(* IEC 61131-3 sources: AI_Prediciton_FInder_Energy_meter/plc/src, 8 files *)

(* ---- U_Word32.st ---- *)
// DUT (UNION) - reinterprets 32 bits as DWORD, REAL or DINT
TYPE U_Word32 :
UNION
    dwRaw : DWORD;
    rReal : REAL;
    diInt : DINT;
END_UNION
END_TYPE

(* ---- GVL_Meter.st ---- *)
// GVL - raw Modbus channels and Modbus TCP input registers
VAR_GLOBAL
    // Finder 7M.24 #1 (Modbus RTU address 2) - mapped in Modbus_Server_COM_Port I/O Mapping
    awFinder1Power      : ARRAY[0..11] OF WORD;  // 32490..32501: Pt, Qt, St, PFt, f, U1 (REAL, high word first)
    awFinder1Current    : ARRAY[0..1] OF WORD;   // 32516..32517: I1 (REAL)
    awFinder1EnergyExp  : ARRAY[0..3] OF WORD;   // 30401..30404: exponents n1..n4 (INT)
    awFinder1EnergyMant : ARRAY[0..7] OF WORD;   // 30406..30413: mantissas n1..n4 (DINT, high word first)
    awFinder1Identity   : ARRAY[0..11] OF WORD;  // 30001..30012: model (0..7) + serial (8..11), ASCII
    awFinder1MaxRegs    : ARRAY[0..0] OF WORD;   // 30099: max registers per request
    // E2-PLC2 (25.11.2026): new channels, existing ones unchanged
    awFinder1Quality    : ARRAY[0..25] OF WORD;  // 32570..32595: angle U1-I1 [0..1], THD I1 [18..19], THD U1 [24..25] (REAL)
    awFinder1Temp       : ARRAY[0..1] OF WORD;   // 32658..32659: internal temperature (REAL, degC)
    awFinder1RunTime    : ARRAY[0..1] OF WORD;   // 32480..32481: run time (REAL, s - type to be confirmed)

    // Modbus TCP server input registers (FC04) - mapped in ModbusTCP_Server_Device I/O Mapping
    awTcpInputRegs      : ARRAY[0..99] OF WORD;
END_VAR

(* ---- FC_PutDword.st ---- *)
// FUNCTION, return type BOOL - writes 32 bits into two registers, high word first
FUNCTION FC_PutDword : BOOL
VAR_IN_OUT
    awRegs : ARRAY[0..99] OF WORD;
END_VAR
VAR_INPUT
    iIndex  : INT;    // index of the first (high) register
    dwValue : DWORD;
END_VAR
// --- code ---
IF (iIndex < 0) OR (iIndex > 98) THEN
    FC_PutDword := FALSE;
    RETURN;
END_IF
awRegs[iIndex]     := DWORD_TO_WORD(SHR(dwValue, 16));
awRegs[iIndex + 1] := DWORD_TO_WORD(dwValue);
FC_PutDword := TRUE;

(* ---- FC_PutReal.st ---- *)
// FUNCTION, return type BOOL - writes REAL (IEEE 754) into two registers, high word first
FUNCTION FC_PutReal : BOOL
VAR_IN_OUT
    awRegs : ARRAY[0..99] OF WORD;
END_VAR
VAR_INPUT
    iIndex : INT;
    rValue : REAL;
END_VAR
VAR
    uConv : U_Word32;
END_VAR
// --- code ---
uConv.rReal := rValue;
FC_PutReal := FC_PutDword(awRegs := awRegs, iIndex := iIndex, dwValue := uConv.dwRaw);

(* ---- FC_WordsToDword.st ---- *)
// FUNCTION, return type DWORD
FUNCTION FC_WordsToDword : DWORD
VAR_INPUT
    wFirst     : WORD;  // register with lower address
    wSecond    : WORD;  // register with higher address
    xSwapWords : BOOL;  // FALSE = first register is the high word (Finder 7M.24, verified 23.11.2026)
END_VAR
// --- code ---
IF xSwapWords THEN
    FC_WordsToDword := SHL(WORD_TO_DWORD(wSecond), 16) OR WORD_TO_DWORD(wFirst);
ELSE
    FC_WordsToDword := SHL(WORD_TO_DWORD(wFirst), 16) OR WORD_TO_DWORD(wSecond);
END_IF

(* ---- FC_WordsToReal.st ---- *)
// FUNCTION, return type REAL
FUNCTION FC_WordsToReal : REAL
VAR_INPUT
    wFirst     : WORD;
    wSecond    : WORD;
    xSwapWords : BOOL;
END_VAR
VAR
    uConv : U_Word32;
END_VAR
// --- code ---
uConv.dwRaw := FC_WordsToDword(wFirst := wFirst, wSecond := wSecond, xSwapWords := xSwapWords);
FC_WordsToReal := uConv.rReal;

(* ---- FB_EnergyMeter.st ---- *)
// FUNCTION_BLOCK - one instance = one Finder 7M.24 meter
FUNCTION_BLOCK FB_EnergyMeter
VAR_INPUT
    xCommError        : BOOL;                   // <device>.xError of the Modbus server (COM) instance
    uiModbusErrorCode : UINT;                   // <device>.byModbusError (MB_ErrorCodes)
    awPower           : ARRAY[0..11] OF WORD;
    awCurrent         : ARRAY[0..1] OF WORD;
    awEnergyExp       : ARRAY[0..3] OF WORD;
    awEnergyMant      : ARRAY[0..7] OF WORD;
    awIdentity        : ARRAY[0..11] OF WORD;
    awQuality         : ARRAY[0..25] OF WORD;   // 32570..32595 (map v2, 25.11.2026)
    awTemp            : ARRAY[0..1] OF WORD;    // 32658..32659
    awRunTime         : ARRAY[0..1] OF WORD;    // 32480..32481
    xSwapWords        : BOOL := FALSE;          // Finder 7M.24: high word first -> FALSE
    tErrorHold        : TIME := T#3S;           // COMM_ERROR is cleared only after this time without any error
END_VAR
VAR_OUTPUT
    rActivePower_W     : REAL;
    rReactivePower_var : REAL;
    rApparentPower_VA  : REAL;
    rPowerFactor       : REAL;
    rFrequency_Hz      : REAL;
    rVoltage_V         : REAL;
    rCurrent_A         : REAL;
    diEnergyImportMant : DINT;   // n1, Wh = mant * 10^exp
    iEnergyImportExp   : INT;
    diEnergyExportMant : DINT;   // n3
    iEnergyExportExp   : INT;
    rEnergyImport_kWh  : REAL;
    rEnergyExport_kWh  : REAL;
    diReactivePosMant  : DINT;   // n2 (energy at Q > 0), varh = mant * 10^exp
    iReactivePosExp    : INT;
    diReactiveNegMant  : DINT;   // n4 (energy at Q < 0)
    iReactiveNegExp    : INT;
    rThdVoltage_pct    : REAL;   // THD U1, 32594
    rThdCurrent_pct    : REAL;   // THD I1, 32588
    rPhaseAngle_deg    : REAL;   // angle U1-I1, 32570 (negative at Q < 0, measured 25.11.2026)
    rTemperature_C     : REAL;   // internal meter temperature, 32658
    rRunTime_s         : REAL;   // meter run time, 32480
    awSerial           : ARRAY[0..3] OF WORD;
    sSerial            : STRING(8);
    uiStatus           : UINT;   // 0 = OK, 1 = COMM_ERROR, 2 = NO_DATA (no answer since start)
    uiErrorCode        : UINT;   // last non-zero MB_ErrorCodes value while not OK, 0 when OK
    uiErrorCount       : UINT;   // number of communication outages since start (wraps at 65535)
    udiDataAge_ms      : UDINT;  // 0 when OK; time since last confirmed OK state otherwise
END_VAR
VAR CONSTANT
    STATUS_OK         : UINT := 0;
    STATUS_COMM_ERROR : UINT := 1;
    STATUS_NO_DATA    : UINT := 2;
END_VAR
VAR
    xErrorSeen       : BOOL;   // at least one raw error since start
    xErrorActive     : BOOL;   // debounced error: raw error within the last tErrorHold
    xErrorActivePrev : BOOL;
    xDataSeen        : BOOL;
    tNow             : TIME;
    tLastOk          : TIME;
    tLastErr         : TIME;
    uiLastErrCode    : UINT;
    uConv            : U_Word32;
    pbySerial        : POINTER TO BYTE;
    i                : INT;
END_VAR
// --- code ---
// 1. Communication status (debounced: xError of the COM device drops between transactions;
//    fixed 23.11.2026 after checklist test 5)
tNow := TIME();
IF xCommError THEN
    xErrorSeen := TRUE;
    tLastErr   := tNow;
    IF uiModbusErrorCode <> 0 THEN
        uiLastErrCode := uiModbusErrorCode;
    END_IF
END_IF

xErrorActive := xErrorSeen AND ((tNow - tLastErr) < tErrorHold);

IF NOT xErrorActive THEN
    tLastOk := tNow;
END_IF
IF xErrorActive AND NOT xErrorActivePrev THEN
    uiErrorCount := uiErrorCount + 1;            // one outage = one count
END_IF
xErrorActivePrev := xErrorActive;

// Meter has answered at least once when the serial number registers are not zero
IF (awIdentity[8] <> 0) OR (awIdentity[9] <> 0) THEN
    xDataSeen := TRUE;
END_IF

IF NOT xDataSeen THEN
    uiStatus      := STATUS_NO_DATA;
    uiErrorCode   := uiLastErrCode;
    udiDataAge_ms := 16#FFFFFFFF;
ELSIF xErrorActive THEN
    uiStatus      := STATUS_COMM_ERROR;
    uiErrorCode   := uiLastErrCode;
    udiDataAge_ms := TIME_TO_UDINT(tNow - tLastOk);
ELSE
    uiStatus      := STATUS_OK;
    uiErrorCode   := 0;
    uiLastErrCode := 0;
    udiDataAge_ms := 0;
END_IF

// 2. Instantaneous values (IEEE 754 block 32490..32501, 32516)
rActivePower_W     := FC_WordsToReal(wFirst := awPower[0],  wSecond := awPower[1],  xSwapWords := xSwapWords);
rReactivePower_var := FC_WordsToReal(wFirst := awPower[2],  wSecond := awPower[3],  xSwapWords := xSwapWords);
rApparentPower_VA  := FC_WordsToReal(wFirst := awPower[4],  wSecond := awPower[5],  xSwapWords := xSwapWords);
rPowerFactor       := FC_WordsToReal(wFirst := awPower[6],  wSecond := awPower[7],  xSwapWords := xSwapWords);
rFrequency_Hz      := FC_WordsToReal(wFirst := awPower[8],  wSecond := awPower[9],  xSwapWords := xSwapWords);
rVoltage_V         := FC_WordsToReal(wFirst := awPower[10], wSecond := awPower[11], xSwapWords := xSwapWords);
rCurrent_A         := FC_WordsToReal(wFirst := awCurrent[0], wSecond := awCurrent[1], xSwapWords := xSwapWords);

// 3. Energy counters: Wh = mantissa * 10^exponent (n1 = import, n3 = export - to confirm on display)
uConv.dwRaw := FC_WordsToDword(wFirst := awEnergyMant[0], wSecond := awEnergyMant[1], xSwapWords := xSwapWords);
diEnergyImportMant := uConv.diInt;
iEnergyImportExp   := WORD_TO_INT(awEnergyExp[0]);

uConv.dwRaw := FC_WordsToDword(wFirst := awEnergyMant[4], wSecond := awEnergyMant[5], xSwapWords := xSwapWords);
diEnergyExportMant := uConv.diInt;
iEnergyExportExp   := WORD_TO_INT(awEnergyExp[2]);

rEnergyImport_kWh := LREAL_TO_REAL(DINT_TO_LREAL(diEnergyImportMant) * EXPT(LREAL#10.0, INT_TO_LREAL(iEnergyImportExp)) / 1000.0);
rEnergyExport_kWh := LREAL_TO_REAL(DINT_TO_LREAL(diEnergyExportMant) * EXPT(LREAL#10.0, INT_TO_LREAL(iEnergyExportExp)) / 1000.0);

// 3b. Reactive energy counters (map v2): n2 = mant[2..3] / exp[1], n4 = mant[6..7] / exp[3]
uConv.dwRaw := FC_WordsToDword(wFirst := awEnergyMant[2], wSecond := awEnergyMant[3], xSwapWords := xSwapWords);
diReactivePosMant := uConv.diInt;
iReactivePosExp   := WORD_TO_INT(awEnergyExp[1]);

uConv.dwRaw := FC_WordsToDword(wFirst := awEnergyMant[6], wSecond := awEnergyMant[7], xSwapWords := xSwapWords);
diReactiveNegMant := uConv.diInt;
iReactiveNegExp   := WORD_TO_INT(awEnergyExp[3]);

// 3c. Power quality, temperature, run time (map v2; values checked online in step PLC-1, 25.11.2026)
rPhaseAngle_deg := FC_WordsToReal(wFirst := awQuality[0],  wSecond := awQuality[1],  xSwapWords := xSwapWords);
rThdCurrent_pct := FC_WordsToReal(wFirst := awQuality[18], wSecond := awQuality[19], xSwapWords := xSwapWords);
rThdVoltage_pct := FC_WordsToReal(wFirst := awQuality[24], wSecond := awQuality[25], xSwapWords := xSwapWords);
rTemperature_C  := FC_WordsToReal(wFirst := awTemp[0],     wSecond := awTemp[1],     xSwapWords := xSwapWords);
rRunTime_s      := FC_WordsToReal(wFirst := awRunTime[0],  wSecond := awRunTime[1],  xSwapWords := xSwapWords);

// 4. Serial number (registers 30009..30012, ASCII, high byte first)
pbySerial := ADR(sSerial);
FOR i := 0 TO 3 DO
    awSerial[i]           := awIdentity[8 + i];
    pbySerial[2 * i]      := WORD_TO_BYTE(SHR(awIdentity[8 + i], 8));
    pbySerial[2 * i + 1]  := WORD_TO_BYTE(awIdentity[8 + i]);
END_FOR
pbySerial[8] := 0;

(* ---- PRG_ModbusTcpMap.st ---- *)
// PROGRAM - reads meter(s) via FB_EnergyMeter and fills Modbus TCP input registers (map v2)
PROGRAM PRG_ModbusTcpMap
VAR CONSTANT
    MAP_VERSION     : WORD := 2;   // v2 since 25.11.2026 (E2-PLC2)
    REG_HEARTBEAT   : INT := 0;   // 0..1  UDINT
    REG_MAP_VERSION : INT := 2;   // 2     UINT
    METER1_BASE     : INT := 10;  // meter block: base .. base+49

    // offsets inside a meter block
    OFS_STATUS      : INT := 0;   // UINT
    OFS_ERROR_CODE  : INT := 1;   // UINT
    OFS_ERROR_COUNT : INT := 2;   // UINT
    OFS_DATA_AGE    : INT := 4;   // UDINT, ms
    OFS_P           : INT := 6;   // REAL, W
    OFS_Q           : INT := 8;   // REAL, var
    OFS_S           : INT := 10;  // REAL, VA
    OFS_PF          : INT := 12;  // REAL
    OFS_F           : INT := 14;  // REAL, Hz
    OFS_U           : INT := 16;  // REAL, V
    OFS_I           : INT := 18;  // REAL, A
    OFS_E_IMP       : INT := 20;  // REAL, kWh
    OFS_E_EXP       : INT := 22;  // REAL, kWh
    OFS_E_IMP_MANT  : INT := 24;  // DINT
    OFS_E_IMP_EXP   : INT := 26;  // INT
    OFS_E_EXP_MANT  : INT := 27;  // DINT
    OFS_E_EXP_EXP   : INT := 29;  // INT
    OFS_SERIAL      : INT := 30;  // 4 x WORD, ASCII
    // map v2
    OFS_Q_POS_MANT  : INT := 34;  // DINT, n2
    OFS_Q_POS_EXP   : INT := 36;  // INT
    OFS_Q_NEG_MANT  : INT := 37;  // DINT, n4
    OFS_Q_NEG_EXP   : INT := 39;  // INT
    OFS_THD_U       : INT := 40;  // REAL, %
    OFS_THD_I       : INT := 42;  // REAL, %
    OFS_ANGLE       : INT := 44;  // REAL, deg
    OFS_TEMP        : INT := 46;  // REAL, degC
    OFS_RUN_TIME    : INT := 48;  // REAL, s
END_VAR
VAR
    udiHeartbeat : UDINT;
    fbMeter1     : FB_EnergyMeter;
    iBase        : INT;
    i            : INT;
END_VAR
// --- code ---
// 1. Meter 1: Finder 7M.24 on COM (Modbus_Server_COM_Port, address 2)
fbMeter1(
    xCommError        := Modbus_Server_COM_Port.xError,
    uiModbusErrorCode := TO_UINT(Modbus_Server_COM_Port.byModbusError),
    awPower           := GVL_Meter.awFinder1Power,
    awCurrent         := GVL_Meter.awFinder1Current,
    awEnergyExp       := GVL_Meter.awFinder1EnergyExp,
    awEnergyMant      := GVL_Meter.awFinder1EnergyMant,
    awIdentity        := GVL_Meter.awFinder1Identity,
    awQuality         := GVL_Meter.awFinder1Quality,
    awTemp            := GVL_Meter.awFinder1Temp,
    awRunTime         := GVL_Meter.awFinder1RunTime,
    xSwapWords        := FALSE);

// 2. Header
udiHeartbeat := udiHeartbeat + 1;
FC_PutDword(awRegs := GVL_Meter.awTcpInputRegs, iIndex := REG_HEARTBEAT, dwValue := UDINT_TO_DWORD(udiHeartbeat));
GVL_Meter.awTcpInputRegs[REG_MAP_VERSION] := MAP_VERSION;

// 3. Meter 1 block
iBase := METER1_BASE;
GVL_Meter.awTcpInputRegs[iBase + OFS_STATUS]      := UINT_TO_WORD(fbMeter1.uiStatus);
GVL_Meter.awTcpInputRegs[iBase + OFS_ERROR_CODE]  := UINT_TO_WORD(fbMeter1.uiErrorCode);
GVL_Meter.awTcpInputRegs[iBase + OFS_ERROR_COUNT] := UINT_TO_WORD(fbMeter1.uiErrorCount);
FC_PutDword(awRegs := GVL_Meter.awTcpInputRegs, iIndex := iBase + OFS_DATA_AGE, dwValue := UDINT_TO_DWORD(fbMeter1.udiDataAge_ms));

FC_PutReal(awRegs := GVL_Meter.awTcpInputRegs, iIndex := iBase + OFS_P,  rValue := fbMeter1.rActivePower_W);
FC_PutReal(awRegs := GVL_Meter.awTcpInputRegs, iIndex := iBase + OFS_Q,  rValue := fbMeter1.rReactivePower_var);
FC_PutReal(awRegs := GVL_Meter.awTcpInputRegs, iIndex := iBase + OFS_S,  rValue := fbMeter1.rApparentPower_VA);
FC_PutReal(awRegs := GVL_Meter.awTcpInputRegs, iIndex := iBase + OFS_PF, rValue := fbMeter1.rPowerFactor);
FC_PutReal(awRegs := GVL_Meter.awTcpInputRegs, iIndex := iBase + OFS_F,  rValue := fbMeter1.rFrequency_Hz);
FC_PutReal(awRegs := GVL_Meter.awTcpInputRegs, iIndex := iBase + OFS_U,  rValue := fbMeter1.rVoltage_V);
FC_PutReal(awRegs := GVL_Meter.awTcpInputRegs, iIndex := iBase + OFS_I,  rValue := fbMeter1.rCurrent_A);
FC_PutReal(awRegs := GVL_Meter.awTcpInputRegs, iIndex := iBase + OFS_E_IMP, rValue := fbMeter1.rEnergyImport_kWh);
FC_PutReal(awRegs := GVL_Meter.awTcpInputRegs, iIndex := iBase + OFS_E_EXP, rValue := fbMeter1.rEnergyExport_kWh);

FC_PutDword(awRegs := GVL_Meter.awTcpInputRegs, iIndex := iBase + OFS_E_IMP_MANT, dwValue := DINT_TO_DWORD(fbMeter1.diEnergyImportMant));
GVL_Meter.awTcpInputRegs[iBase + OFS_E_IMP_EXP] := INT_TO_WORD(fbMeter1.iEnergyImportExp);
FC_PutDword(awRegs := GVL_Meter.awTcpInputRegs, iIndex := iBase + OFS_E_EXP_MANT, dwValue := DINT_TO_DWORD(fbMeter1.diEnergyExportMant));
GVL_Meter.awTcpInputRegs[iBase + OFS_E_EXP_EXP] := INT_TO_WORD(fbMeter1.iEnergyExportExp);

FOR i := 0 TO 3 DO
    GVL_Meter.awTcpInputRegs[iBase + OFS_SERIAL + i] := fbMeter1.awSerial[i];
END_FOR

// 4. Map v2: registers 44..59 (offsets 34..49)
FC_PutDword(awRegs := GVL_Meter.awTcpInputRegs, iIndex := iBase + OFS_Q_POS_MANT, dwValue := DINT_TO_DWORD(fbMeter1.diReactivePosMant));
GVL_Meter.awTcpInputRegs[iBase + OFS_Q_POS_EXP] := INT_TO_WORD(fbMeter1.iReactivePosExp);
FC_PutDword(awRegs := GVL_Meter.awTcpInputRegs, iIndex := iBase + OFS_Q_NEG_MANT, dwValue := DINT_TO_DWORD(fbMeter1.diReactiveNegMant));
GVL_Meter.awTcpInputRegs[iBase + OFS_Q_NEG_EXP] := INT_TO_WORD(fbMeter1.iReactiveNegExp);
FC_PutReal(awRegs := GVL_Meter.awTcpInputRegs, iIndex := iBase + OFS_THD_U,    rValue := fbMeter1.rThdVoltage_pct);
FC_PutReal(awRegs := GVL_Meter.awTcpInputRegs, iIndex := iBase + OFS_THD_I,    rValue := fbMeter1.rThdCurrent_pct);
FC_PutReal(awRegs := GVL_Meter.awTcpInputRegs, iIndex := iBase + OFS_ANGLE,    rValue := fbMeter1.rPhaseAngle_deg);
FC_PutReal(awRegs := GVL_Meter.awTcpInputRegs, iIndex := iBase + OFS_TEMP,     rValue := fbMeter1.rTemperature_C);
FC_PutReal(awRegs := GVL_Meter.awTcpInputRegs, iIndex := iBase + OFS_RUN_TIME, rValue := fbMeter1.rRunTime_s);
